            num nSigValue = 1
        pointRx pPointRx[2] = {x=490.110293, y=-600.305611, z=568.056156, rx=-6.599443, ry=-2.68541, rz=28.351195, shoulder=lefty, elbow=enegative, wrist=wpositive}
        string sID
      [48]
        bool bMarked
        jointRx jJointRx = {j1=-87.551314, j2=145.129335, j3=-83.085728, j4=182.11845, j5=63.691243, j6=-64.966658}
        pointRx pInter
        paraItem pParaItem
          [0]
            bool bSafePoint
            ifItem iIfItem
              [0]
                bool bANDOR[2]
                num nSigIndex[3]
                num nSigType[3]
                num nValue[3]
            mdesc mMdesc
            num nActionIndex = 42
            num nDelay
            num nMoveType = 1
            num nPercentage
            num nSigValue = 1
        pointRx pPointRx[2] = {x=61.349727, y=-652.129552, z=350.0734551, rx=-1.549449, ry=-1.96692, rz=28.421736, shoulder=lefty, elbow=enegative, wrist=wpositive}
        string sID
    string sID
  [Position6_point_blow]
    num nFrameIndex
    num nMoveID
    num nToolIndex
    pointItem pPointItem[64]
      [0]
        bool bMarked
        jointRx jJointRx
        pointRx pInter
        paraItem pParaItem
          [0]
            bool bSafePoint
            ifItem iIfItem
              [0]
                bool bANDOR[2]
                num nSigIndex[3]
                num nSigType[3]
                num nValue[3]
            mdesc mMdesc
            num nActionIndex = 43
            num nDelay
            num nMoveType = 4
            num nPercentage
            num nSigValue = 1
        pointRx pPointRx[2]
        string sID
      [1]
        bool bMarked
        jointRx jJointRx = {j1=-87.550712, j2=145.128314, j3=-83.0892365, j4=182.11811, j5=63.690987, j6=-64.966608}
        pointRx pInter
        paraItem pParaItem
          [0]
            bool bSafePoint
            ifItem iIfItem
              [0]
                bool bANDOR[2]
                num nSigIndex[3]
                num nSigType[3]
                num nValue[3]
            mdesc mMdesc
            num nActionIndex = 42
            num nDelay
            num nMoveType = 1
            num nPercentage
            num nSigValue = 1
        pointRx pPointRx[2] = {x=61.357264, y=-652.082, z=350.106484, rx=-1.553715, ry=-1.966811, rz=28.422241, shoulder=lefty, elbow=enegative, wrist=wpositive}
        string sID
      [2]
        bool bMarked
        jointRx jJointRx = {j1=-58.982134, j2=104.832128, j3=-61.565333, j4=183.343645, j5=42.668286, j6=-33.606181}
        pointRx pInter
        paraItem pParaItem
          [0]
            bool bSafePoint
            ifItem iIfItem
              [0]
                bool bANDOR[2]
                num nSigIndex[3]
                num nSigType[3]
                num nValue[3]
            mdesc mMdesc
            num nActionIndex = 42
            num nDelay
            num nMoveType = 1
            num nPercentage
            num nSigValue = 1
        pointRx pPointRx[2] = {x=416.397495, y=-633.838238, z=700.254781, rx=1.722211, ry=-1.608013, rz=89.88289, shoulder=lefty, elbow=enegative, wrist=wpositive}
        string sID
      [3]
        bool bMarked
        jointRx jJointRx = {j1=-62.332645, j2=107.50753, j3=-68.132801, j4=183.562396, j5=38.651057, j6=-30.577163}
        pointRx pInter
        paraItem pParaItem
          [0]
            bool bSafePoint
            ifItem iIfItem
              [0]
                bool bANDOR[2]
                num nSigIndex[3]
                num nSigType[3]
                num nValue[3]
            mdesc mMdesc
            num nActionIndex = 42
            num nDelay
            num nMoveType = 1
            num nPercentage
            num nSigValue = 1
        pointRx pPointRx[2] = {x=366.85786, y=-633.838275, z=700.254798, rx=1.721666, ry=-1.608681, rz=89.88277, shoulder=lefty, elbow=enegative, wrist=wpositive}
        string sID
      [4]
        bool bMarked
        jointRx jJointRx = {j1=-67.0327916, j2=110.2281, j3=-75.107293, j4=183.830258, j5=34.223084, j6=-26.259259}
        pointRx pInter
        paraItem pParaItem
          [0]
            bool bSafePoint
            ifItem iIfItem
              [0]
                bool bANDOR[2]
                num nSigIndex[3]
                num nSigType[3]
                num nValue[3]
            mdesc mMdesc
            num nActionIndex = 42
            num nDelay
            num nMoveType = 1
            num nPercentage
            num nSigValue = 1
        pointRx pPointRx[2] = {x=302.522929, y=-633.83826, z=700.254794, rx=1.721622, ry=-1.608914, rz=89.882692, shoulder=lefty, elbow=enegative, wrist=wpositive}
        string sID
      [5]
        bool bMarked
        jointRx jJointRx = {j1=-71.633736, j2=112.694899, j3=-81.788319, j4=184.160101, j5=29.845031, j6=-22.0972061}
        pointRx pInter
        paraItem pParaItem
          [0]
            bool bSafePoint
            ifItem iIfItem
              [0]
                bool bANDOR[2]
                num nSigIndex[3]
                num nSigType[3]
                num nValue[3]
            mdesc mMdesc
            num nActionIndex = 42
            num nDelay
            num nMoveType = 1
            num nPercentage
            num nSigValue = 1
        pointRx pPointRx[2] = {x=241.500206, y=-626.00943449, z=700.254792, rx=1.721289, ry=-1.608551, rz=89.882813, shoulder=lefty, elbow=enegative, wrist=wpositive}
        string sID
      [6]
        bool bMarked
        jointRx jJointRx = {j1=-65.27374, j2=114.413405, j3=-86.726434, j4=184.827216, j5=26.876761, j6=-29.158228}
        pointRx pInter
        paraItem pParaItem
          [0]
            bool bSafePoint
            ifItem iIfItem
              [0]
                bool bANDOR[2]
                num nSigIndex[3]
                num nSigType[3]
                num nValue[3]
            mdesc mMdesc
            num nActionIndex = 42
            num nDelay
            num nMoveType = 1
            num nPercentage
            num nSigValue = 1
        pointRx pPointRx[2] = {x=296.78184, y=-570.410131, z=700.254763, rx=1.722456, ry=-1.607129, rz=89.88308, shoulder=lefty, elbow=enegative, wrist=wpositive}
        string sID
      [7]
        bool bMarked
        jointRx jJointRx = {j1=-60.709616, j2=114.554511, j3=-87.145192, j4=184.986355, j5=26.782513, j6=-33.871303}
        pointRx pInter
        paraItem pParaItem
          [0]
            bool bSafePoint
            ifItem iIfItem
              [0]
                bool bANDOR[2]
                num nSigIndex[3]
                num nSigType[3]
                num nValue[3]
            mdesc mMdesc
            num nActionIndex = 42
            num nDelay
            num nMoveType = 1
            num nPercentage
            num nSigValue = 1
        pointRx pPointRx[2] = {x=338.875527, y=-541.934118, z=700.254791, rx=1.721113, ry=-1.608268, rz=89.882966, shoulder=lefty, elbow=enegative, wrist=wpositive}
        string sID
      [8]
        bool bMarked
        jointRx jJointRx = {j1=-66.643474, j2=118.657481, j3=-100.787497, j4=187.380827, j5=17.0599953, j6=-30.539636}
        pointRx pInter
        paraItem pParaItem
          [0]
            bool bSafePoint
            ifItem iIfItem
              [0]
                bool bANDOR[2]
                num nSigIndex[3]
                num nSigType[3]
                num nValue[3]
            mdesc mMdesc
            num nActionIndex = 42
            num nDelay
            num nMoveType = 1
            num nPercentage
            num nSigValue = 1
        pointRx pPointRx[2] = {x=251.241513, y=-503.208169, z=700.254788, rx=1.722301, ry=-1.608953, rz=89.882703, shoulder=lefty, elbow=enegative, wrist=wpositive}
        string sID
      [9]
        bool bMarked
        jointRx jJointRx = {j1=-65.0394334, j2=119.495527, j3=-104.191107, j4=188.704216, j5=14.582841, j6=-33.512784}
        pointRx pInter
        paraItem pParaItem
          [0]
            bool bSafePoint
            ifItem iIfItem
              [0]
                bool bANDOR[2]
                num nSigIndex[3]
                num nSigType[3]
                num nValue[3]
            mdesc mMdesc
            num nActionIndex = 42
            num nDelay
            num nMoveType = 1
            num nPercentage
            num nSigValue = 1
        pointRx pPointRx[2] = {x=255.846551, y=-476.313024, z=700.254767, rx=1.721654, ry=-1.607307, rz=89.883015, shoulder=lefty, elbow=enegative, wrist=wpositive}
        string sID
      [10]
        bool bMarked
        jointRx jJointRx = {j1=-71.0596735, j2=121.00750191, j3=-111.877772, j4=194.578806, j5=8.286602, j6=-33.494479}
        pointRx pInter
        paraItem pParaItem
          [0]
            bool bSafePoint
            ifItem iIfItem
              [0]
                bool bANDOR[2]
                num nSigIndex[3]
                num nSigType[3]
                num nValue[3]
            mdesc mMdesc
            num nActionIndex = 42
            num nDelay
            num nMoveType = 1
            num nPercentage
            num nSigValue = 1
        pointRx pPointRx[2] = {x=189.620191, y=-454.405925, z=700.254767, rx=1.721353, ry=-1.607377, rz=89.882905, shoulder=lefty, elbow=enegative, wrist=wpositive}
        string sID
      [11]
        bool bMarked
        jointRx jJointRx = {j1=-74.809464, j2=121.0382904, j3=-112.0769955, j4=194.59856, j5=7.974501, j6=-29.773551}
        pointRx pInter
        paraItem pParaItem
          [0]
            bool bSafePoint
            ifItem iIfItem
              [0]
                bool bANDOR[2]
                num nSigIndex[3]
                num nSigType[3]
                num nValue[3]
            mdesc mMdesc
            num nActionIndex = 42
            num nDelay
            num nMoveType = 1
            num nPercentage
            num nSigValue = 1
        pointRx pPointRx[2] = {x=160.082647, y=-465.491863, z=700.254784, rx=1.722803, ry=-1.608682, rz=89.882806, shoulder=lefty, elbow=enegative, wrist=wpositive}
        string sID
      [12]
        bool bMarked
        jointRx jJointRx = {j1=-76.815291, j2=120.680634, j3=-109.926019, j4=191.777648, j5=9.643692, j6=-24.919524}
        pointRx pInter
        paraItem pParaItem
          [0]
            bool bSafePoint
            ifItem iIfItem
              [0]
                bool bANDOR[2]
                num nSigIndex[3]
                num nSigType[3]
                num nValue[3]
            mdesc mMdesc
            num nActionIndex = 42
            num nDelay
            num nMoveType = 1
            num nPercentage
            num nSigValue = 1
        pointRx pPointRx[2] = {x=147.50556, y=-485.393693, z=700.254789, rx=1.722658, ry=-1.609045, rz=89.882735, shoulder=lefty, elbow=enegative, wrist=wpositive}
        string sID
      [13]
        bool bMarked
        jointRx jJointRx = {j1=-80.979539, j2=121.627826, j3=-116.887787, j4=209.4559, j5=3.779386, j6=-38.540773}
        pointRx pInter
        paraItem pParaItem
          [0]
            bool bSafePoint
            ifItem iIfItem
              [0]
                bool bANDOR[2]
                num nSigIndex[3]
                num nSigType[3]
                num nValue[3]
            mdesc mMdesc
            num nActionIndex = 42
            num nDelay
            num nMoveType = 1
            num nPercentage
            num nSigValue = 1
        pointRx pPointRx[2] = {x=105.438294, y=-448.641412, z=700.254346, rx=1.721348, ry=-1.60753, rz=89.882882, shoulder=lefty, elbow=enegative, wrist=wpositive}
        string sID
      [14]
        bool bMarked
        jointRx jJointRx = {j1=-97.0735787, j2=120.583034, j3=-109.386983, j4=169.0121648, j5=9.967554, j6=107.0502076}
        pointRx pInter
        paraItem pParaItem
          [0]
            bool bSafePoint
            ifItem iIfItem
              [0]
                bool bANDOR[2]
                num nSigIndex[3]
                num nSigType[3]
                num nValue[3]
            mdesc mMdesc
            num nActionIndex = 42
            num nDelay
            num nMoveType = 1
            num nPercentage
            num nSigValue = 1
        pointRx pPointRx[2] = {x=3.102788, y=-514.97816, z=700.254373, rx=1.629756, ry=1.702884, rz=179.149702, shoulder=lefty, elbow=enegative, wrist=wpositive}
        string sID
      [15]
        bool bMarked
        jointRx jJointRx = {j1=-98.785966, j2=121.589944, j3=-116.474742, j4=152.822693, j5=4.230949, j6=125.0509123}
        pointRx pInter
        paraItem pParaItem
          [0]
            bool bSafePoint
            ifItem iIfItem
              [0]
                bool bANDOR[2]
                num nSigIndex[3]
                num nSigType[3]
                num nValue[3]
            mdesc mMdesc
            num nActionIndex = 42
            num nDelay
            num nMoveType = 1
            num nPercentage
            num nSigValue = 1
        pointRx pPointRx[2] = {x=-4.455751, y=-466.481228, z=700.254288, rx=1.629056, ry=1.702249, rz=179.149669, shoulder=lefty, elbow=enegative, wrist=wpositive}
        string sID
      [16]
        bool bMarked
        jointRx jJointRx = {j1=-102.289362, j2=121.662055, j3=-117.287244, j4=147.396601, j5=3.732456, j6=133.989908}
        pointRx pInter
        paraItem pParaItem
          [0]
            bool bSafePoint
            ifItem iIfItem
              [0]
                bool bANDOR[2]
                num nSigIndex[3]
                num nSigType[3]
                num nValue[3]
            mdesc mMdesc
            num nActionIndex = 42
            num nDelay
            num nMoveType = 1
            num nPercentage
            num nSigValue = 1
        pointRx pPointRx[2] = {x=-30.830703, y=-458.833227, z=700.253116, rx=1.628925, ry=1.702444, rz=179.149706, shoulder=lefty, elbow=enegative, wrist=wpositive}
        string sID
      [17]
        bool bMarked
        jointRx jJointRx = {j1=-97.596795, j2=121.636094, j3=-116.996972, j4=154.0724475, j5=5.372504, j6=163.484863}
        pointRx pInter
        paraItem pParaItem
          [0]
            bool bSafePoint
            ifItem iIfItem
              [0]
                bool bANDOR[2]
                num nSigIndex[3]
                num nSigType[3]
                num nValue[3]
            mdesc mMdesc
            num nActionIndex = 42
            num nDelay
            num nMoveType = 1
            num nPercentage
            num nSigValue = 1
        pointRx pPointRx[2] = {x=11.0855283, y=-449.928798, z=700.263578, rx=0.116735, ry=2.351476, rz=-139.946822, shoulder=lefty, elbow=enegative, wrist=wpositive}
        string sID
      [18]
        bool bMarked
        jointRx jJointRx = {j1=-93.435678, j2=120.973902, j3=-111.67187, j4=165.758899, j5=9.616057, j6=147.540776}
        pointRx pInter
        paraItem pParaItem
          [0]
            bool bSafePoint
            ifItem iIfItem
              [0]
                bool bANDOR[2]
                num nSigIndex[3]
                num nSigType[3]
                num nValue[3]
            mdesc mMdesc
            num nActionIndex = 42
            num nDelay
            num nMoveType = 1
            num nPercentage
            num nSigValue = 1
        pointRx pPointRx[2] = {x=41.481677, y=-486.244692, z=700.26363, rx=0.117474, ry=2.35234, rz=-139.946783, shoulder=lefty, elbow=enegative, wrist=wpositive}
        string sID
      [19]
        bool bMarked
        jointRx jJointRx = {j1=-87.514361, j2=121.638618, j3=-117.0243701, j4=151.901605, j5=4.980778, j6=155.573887}
        pointRx pInter
        paraItem pParaItem
          [0]
            bool bSafePoint
            ifItem iIfItem
              [0]
                bool bANDOR[2]
                num nSigIndex[3]
                num nSigType[3]
                num nValue[3]
            mdesc mMdesc
            num nActionIndex = 42
            num nDelay
            num nMoveType = 1
            num nPercentage
            num nSigValue = 1
        pointRx pPointRx[2] = {x=89.805675, y=-444.448305, z=700.262762, rx=0.116151, ry=2.350833, rz=-139.946826, shoulder=lefty, elbow=enegative, wrist=wpositive}
        string sID
      [20]
        bool bMarked
        jointRx jJointRx = {j1=-85.538373, j2=121.159338, j3=-112.89672, j4=163.596021, j5=8.296682, j6=141.829296}
        pointRx pInter
        paraItem pParaItem
          [0]
            bool bSafePoint
            ifItem iIfItem
              [0]
                bool bANDOR[2]
                num nSigIndex[3]
                num nSigType[3]
                num nValue[3]
            mdesc mMdesc
            num nActionIndex = 42
            num nDelay
            num nMoveType = 1
            num nPercentage
            num nSigValue = 1
        pointRx pPointRx[2] = {x=107.297774, y=-470.450865, z=700.262819, rx=0.116544, ry=2.351714, rz=-139.94676, shoulder=lefty, elbow=enegative, wrist=wpositive}
        string sID
      [21]
        bool bMarked
        jointRx jJointRx = {j1=-80.389938, j2=121.305327, j3=-113.961147, j4=161.375696, j5=7.211507, j6=138.92232}
        pointRx pInter
        paraItem pParaItem
          [0]
            bool bSafePoint
            ifItem iIfItem
              [0]
                bool bANDOR[2]
                num nSigIndex[3]
                num nSigType[3]
                num nValue[3]
            mdesc mMdesc
            num nActionIndex = 42
            num nDelay
            num nMoveType = 1
            num nPercentage
            num nSigValue = 1
        pointRx pPointRx[2] = {x=147.836969, y=-453.554332, z=700.262491, rx=0.115759, ry=2.349936, rz=-139.946858, shoulder=lefty, elbow=enegative, wrist=wpositive}
        string sID
      [22]
        bool bMarked
        jointRx jJointRx = {j1=-74.160542, j2=121.48868, j3=-115.480429, j4=163.296331, j5=4.15176, j6=89.975533}
        pointRx pInter
        paraItem pParaItem
          [0]
            bool bSafePoint
            ifItem iIfItem
              [0]
                bool bANDOR[2]
                num nSigIndex[3]
                num nSigType[3]
                num nValue[3]
            mdesc mMdesc
            num nActionIndex = 42
            num nDelay
            num nMoveType = 1
            num nPercentage
            num nSigValue = 1
        pointRx pPointRx[2] = {x=187.654652, y=-440.110471, z=700.252779, rx=1.628669, ry=1.701382, rz=179.149675, shoulder=lefty, elbow=enegative, wrist=wpositive}
        string sID
      [23]
        bool bMarked
        jointRx jJointRx = {j1=-69.509661, j2=119.265921, j3=-103.220112, j4=175.749132, j5=13.961301, j6=72.790426}
        pointRx pInter
        paraItem pParaItem
          [0]
            bool bSafePoint
            ifItem iIfItem
              [0]
                bool bANDOR[2]
                num nSigIndex[3]
                num nSigType[3]
                num nValue[3]
            mdesc mMdesc
            num nActionIndex = 42
            num nDelay
            num nMoveType = 1
            num nPercentage
            num nSigValue = 1
        pointRx pPointRx[2] = {x=250.0960558, y=-500.875002, z=700.252775, rx=1.628687, ry=1.702386, rz=179.149806, shoulder=lefty, elbow=enegative, wrist=wpositive}
        string sID
      [24]
        bool bMarked
        jointRx jJointRx = {j1=-65.451313, j2=120.0346612, j3=-106.615882, j4=175.540521, j5=11.264344, j6=68.982362}
        pointRx pInter
        paraItem pParaItem
          [0]
            bool bSafePoint
            ifItem iIfItem
              [0]
                bool bANDOR[2]
                num nSigIndex[3]
                num nSigType[3]
                num nValue[3]
            mdesc mMdesc
            num nActionIndex = 42
            num nDelay
            num nMoveType = 1
            num nPercentage
            num nSigValue = 1
        pointRx pPointRx[2] = {x=274.930404, y=-463.298611, z=700.25277, rx=1.6286, ry=1.700384, rz=179.149585, shoulder=lefty, elbow=enegative, wrist=wpositive}
        string sID
      [25]
        bool bMarked
        jointRx jJointRx = {j1=-63.0913911, j2=120.463088, j3=-108.745441, j4=175.274971, j5=9.527094, j6=66.910352}
        pointRx pInter
        paraItem pParaItem
          [0]
            bool bSafePoint
            ifItem iIfItem
              [0]
                bool bANDOR[2]
                num nSigIndex[3]
                num nSigType[3]
                num nValue[3]
            mdesc mMdesc
            num nActionIndex = 42
            num nDelay
            num nMoveType = 1
            num nPercentage
            num nSigValue = 1
        pointRx pPointRx[2] = {x=286.920288, y=-439.796835, z=700.252783, rx=1.628449, ry=1.702261, rz=179.149771, shoulder=lefty, elbow=enegative, wrist=wpositive}
        string sID
      [26]
        bool bMarked
        jointRx jJointRx = {j1=-60.107122, j2=120.743514, j3=-110.280684, j4=175.353325, j5=8.229554, j6=63.86699}
        pointRx pInter
        paraItem pParaItem
          [0]
            bool bSafePoint
            ifItem iIfItem
              [0]
                bool bANDOR[2]
                num nSigIndex[3]
                num nSigType[3]
                num nValue[3]
            mdesc mMdesc
            num nActionIndex = 42
            num nDelay
            num nMoveType = 1
            num nPercentage
            num nSigValue = 1
        pointRx pPointRx[2] = {x=303.628134, y=-416.218815, z=700.252788, rx=1.628466, ry=1.702202, rz=179.149747, shoulder=lefty, elbow=enegative, wrist=wpositive}
        string sID
      [27]
        bool bMarked
        jointRx jJointRx = {j1=-63.992151, j2=118.544695, j3=-100.353777, j4=177.0428516, j5=16.00047448, j6=65.992969}
        pointRx pInter
        paraItem pParaItem
          [0]
            bool bSafePoint
            ifItem iIfItem
              [0]
                bool bANDOR[2]
                num nSigIndex[3]
                num nSigType[3]
                num nValue[3]
            mdesc mMdesc
            num nActionIndex = 42
            num nDelay
            num nMoveType = 1
            num nPercentage
            num nSigValue = 1
        pointRx pPointRx[2] = {x=303.593559, y=-492.00120121, z=700.25275, rx=1.629773, ry=1.701529, rz=179.149557, shoulder=lefty, elbow=enegative, wrist=wpositive}
        string sID
      [28]
        bool bMarked
        jointRx jJointRx = {j1=-65.604658, j2=115.34522, j3=-89.535997, j4=177.811149, j5=23.638027, j6=66.767236}
        pointRx pInter
        paraItem pParaItem
          [0]
            bool bSafePoint
            ifItem iIfItem
              [0]
                bool bANDOR[2]
                num nSigIndex[3]
                num nSigType[3]
                num nValue[3]
            mdesc mMdesc
            num nActionIndex = 42
            num nDelay
            num nMoveType = 1
            num nPercentage
            num nSigValue = 1
        pointRx pPointRx[2] = {x=316.105522, y=-557.406438, z=700.252765, rx=1.629152, ry=1.702122, rz=179.149764, shoulder=lefty, elbow=enegative, wrist=wpositive}
        string sID
      [29]
        bool bMarked
        jointRx jJointRx = {j1=-68.955824, j2=108.932967, j3=-71.74331, j4=178.253914, j5=35.0703752, j6=69.540198}
        pointRx pInter
        paraItem pParaItem
          [0]
            bool bSafePoint
            ifItem iIfItem
              [0]
                bool bANDOR[2]
                num nSigIndex[3]
                num nSigType[3]
                num nValue[3]
            mdesc mMdesc
            num nActionIndex = 42
            num nDelay
            num nMoveType = 1
            num nPercentage
            num nSigValue = 1
        pointRx pPointRx[2] = {x=316.0702808, y=-657.877777, z=700.252731, rx=1.629581, ry=1.701668, rz=179.149612, shoulder=lefty, elbow=enegative, wrist=wpositive}
        string sID
      [30]
        bool bMarked
        jointRx jJointRx = {j1=-63.428303, j2=105.599126, j3=-63.42748, j4=178.764025, j5=39.960548, j6=63.523315}
        pointRx pInter
        paraItem pParaItem
          [0]
            bool bSafePoint
            ifItem iIfItem
              [0]
                bool bANDOR[2]
                num nSigIndex[3]
                num nSigType[3]
                num nValue[3]
            mdesc mMdesc
            num nActionIndex = 42
            num nDelay
            num nMoveType = 1
            num nPercentage
            num nSigValue = 1
        pointRx pPointRx[2] = {x=392.672125, y=-657.853849, z=700.276087, rx=1.628612, ry=1.701821, rz=179.138765, shoulder=lefty, elbow=enegative, wrist=wpositive}
        string sID
      [31]
        bool bMarked
        jointRx jJointRx = {j1=-64.321332, j2=88.690196, j3=-45.113442, j4=178.747654, j5=41.378269, j6=64.407958}
        pointRx pInter
        paraItem pParaItem
          [0]
            bool bSafePoint
            ifItem iIfItem
              [0]
                bool bANDOR[2]
                num nSigIndex[3]
                num nSigType[3]
                num nValue[3]
            mdesc mMdesc
            num nActionIndex = 42
            num nDelay
            num nMoveType = 1
            num nPercentage
            num nSigValue = 1
        pointRx pPointRx[2] = {x=392.636913, y=-684.559631, z=817.184286, rx=1.629027, ry=1.701529, rz=179.138589, shoulder=lefty, elbow=enegative, wrist=wpositive}
        string sID
      [32]
        bool bMarked
        jointRx jJointRx = {j1=-64.968443, j2=76.908071, j3=-27.68217, j4=178.834761, j5=47.0360379, j6=64.909112}
        pointRx pInter
        paraItem pParaItem
          [0]
            bool bSafePoint
            ifItem iIfItem
              [0]
                bool bANDOR[2]
                num nSigIndex[3]
                num nSigType[3]
                num nValue[3]
            mdesc mMdesc
            num nActionIndex = 42
            num nDelay
            num nMoveType = 1
            num nPercentage
            num nSigValue = 1
        pointRx pPointRx[2] = {x=392.63674, y=-705.0468714, z=873.404329, rx=1.628998, ry=1.701548, rz=179.138605, shoulder=lefty, elbow=enegative, wrist=wpositive}
        string sID
      [33]
        bool bMarked
        jointRx jJointRx = {j1=-62.336449, j2=89.481455, j3=-54.547425, j4=178.610325, j5=32.711346, j6=62.654003}
        pointRx pInter
        paraItem pParaItem
          [0]
            bool bSafePoint
            ifItem iIfItem
              [0]
                bool bANDOR[2]
                num nSigIndex[3]
                num nSigType[3]
                num nValue[3]
            mdesc mMdesc
            num nActionIndex = 42
            num nDelay
            num nMoveType = 1
            num nPercentage
            num nSigValue = 1
        pointRx pPointRx[2] = {x=392.637106, y=-627.212597, z=851.844705, rx=1.627027, ry=1.700481, rz=179.138679, shoulder=lefty, elbow=enegative, wrist=wpositive}
        string sID
      [34]
        bool bMarked
        jointRx jJointRx = {j1=-60.214263, j2=94.794241, j3=-66.773415, j4=178.463697, j5=25.772301, j6=60.747514}
        pointRx pInter
        paraItem pParaItem
          [0]
            bool bSafePoint
            ifItem iIfItem
              [0]
                bool bANDOR[2]
                num nSigIndex[3]
                num nSigType[3]
                num nValue[3]
            mdesc mMdesc
            num nActionIndex = 42
            num nDelay
            num nMoveType = 1
            num nPercentage
            num nSigValue = 1
        pointRx pPointRx[2] = {x=392.637091, y=-573.593172, z=839.237969, rx=1.626982, ry=1.700524, rz=179.13871, shoulder=lefty, elbow=enegative, wrist=wpositive}
        string sID
      [35]
        bool bMarked
        jointRx jJointRx = {j1=-55.995459, j2=94.871223, j3=-77.350718, j4=178.0932115, j5=15.228667, j6=56.988296}
        pointRx pInter
        paraItem pParaItem
          [0]
            bool bSafePoint
            ifItem iIfItem
              [0]
                bool bANDOR[2]
                num nSigIndex[3]
                num nSigType[3]
                num nValue[3]
            mdesc mMdesc
            num nActionIndex = 42
            num nDelay
            num nMoveType = 1
            num nPercentage
            num nSigValue = 1
        pointRx pPointRx[2] = {x=392.637078, y=-484.790879, z=868.772586, rx=1.626877, ry=1.701216, rz=179.138854, shoulder=lefty, elbow=enegative, wrist=wpositive}
        string sID
      [36]
        bool bMarked
        jointRx jJointRx = {j1=-58.229299, j2=114.285829, j3=-86.304494, j4=178.642261, j5=25.707127, j6=58.603666}
        pointRx pInter
        paraItem pParaItem
          [0]
            bool bSafePoint
            ifItem iIfItem
              [0]
                bool bANDOR[2]
                num nSigIndex[3]
                num nSigType[3]
                num nValue[3]
            mdesc mMdesc
            num nActionIndex = 42
            num nDelay
            num nMoveType = 1
            num nPercentage
            num nSigValue = 1
        pointRx pPointRx[2] = {x=392.637007, y=-529.258957, z=700.0975269, rx=1.629049, ry=1.701252, rz=179.138503, shoulder=lefty, elbow=enegative, wrist=wpositive}
        string sID
      [37]
        bool bMarked
        jointRx jJointRx = {j1=-82.703196, j2=116.122044, j3=-91.853722, j4=179.533458, j5=22.561363, j6=-8.781235}
        pointRx pInter
        paraItem pParaItem
          [0]
            bool bSafePoint
            ifItem iIfItem
              [0]
                bool bANDOR[2]
                num nSigIndex[3]
                num nSigType[3]
                num nValue[3]
            mdesc mMdesc
            num nActionIndex = 42
            num nDelay
            num nMoveType = 1
            num nPercentage
            num nSigValue = 1
        pointRx pPointRx[2] = {x=130.0386713, y=-609.589422, z=700.0975633, rx=1.671086, ry=0.394403, rz=88.0816451, shoulder=lefty, elbow=enegative, wrist=wpositive}
        string sID
      [38]
        bool bMarked
        jointRx jJointRx = {j1=-82.0614145, j2=118.602251, j3=-100.420616, j4=179.303357, j5=16.477589, j6=-7.920976}
        pointRx pInter
        paraItem pParaItem
          [0]
            bool bSafePoint
            ifItem iIfItem
              [0]
                bool bANDOR[2]
                num nSigIndex[3]
                num nSigType[3]
                num nValue[3]
            mdesc mMdesc
            num nActionIndex = 42
            num nDelay
            num nMoveType = 1
            num nPercentage
            num nSigValue = 1
        pointRx pPointRx[2] = {x=130.0386769, y=-558.013851, z=700.0975609, rx=1.661587, ry=0.431173, rz=89.346263, shoulder=lefty, elbow=enegative, wrist=wpositive}
        string sID
      [39]
        bool bMarked
        jointRx jJointRx = {j1=-90.0104561, j2=120.70672, j3=-109.816065, j4=177.317534, j5=9.238811, j6=2.005015}
        pointRx pInter
        paraItem pParaItem
          [0]
            bool bSafePoint
            ifItem iIfItem
              [0]
                bool bANDOR[2]
                num nSigIndex[3]
                num nSigType[3]
                num nValue[3]
            mdesc mMdesc
            num nActionIndex = 42
            num nDelay
            num nMoveType = 1
            num nPercentage
            num nSigValue = 1
        pointRx pPointRx[2] = {x=53.663817, y=-510.218495, z=700.0975573, rx=1.661871, ry=0.430213, rz=89.346845, shoulder=lefty, elbow=enegative, wrist=wpositive}
        string sID
      [40]
        bool bMarked
        jointRx jJointRx = {j1=-98.300868, j2=121.852736, j3=-119.389976, j4=142.928524, j5=1.104688, j6=44.711227}
        pointRx pInter
        paraItem pParaItem
          [0]
            bool bSafePoint
            ifItem iIfItem
              [0]
                bool bANDOR[2]
                num nSigIndex[3]
                num nSigType[3]
                num nValue[3]
            mdesc mMdesc
            num nActionIndex = 42
            num nDelay
            num nMoveType = 1
            num nPercentage
            num nSigValue = 1
        pointRx pPointRx[2] = {x=-8.738518, y=-446.473036, z=700.0947095, rx=1.660849, ry=0.430654, rz=89.346953, shoulder=lefty, elbow=enegative, wrist=wpositive}
        string sID
      [41]
        bool bMarked
        jointRx jJointRx = {j1=-101.944431, j2=121.840245, j3=-119.156799, j4=146.219817, j5=1.37852, j6=45.0598803}
        pointRx pInter
        paraItem pParaItem
          [0]
            bool bSafePoint
            ifItem iIfItem
              [0]
                bool bANDOR[2]
                num nSigIndex[3]
                num nSigType[3]
                num nValue[3]
            mdesc mMdesc
            num nActionIndex = 42
            num nDelay
            num nMoveType = 1
            num nPercentage
            num nSigValue = 1
        pointRx pPointRx[2] = {x=-36.505296, y=-446.471107, z=700.0993486, rx=1.662873, ry=0.431649, rz=89.346951, shoulder=lefty, elbow=enegative, wrist=wpositive}
        string sID
      [42]
        bool bMarked
        jointRx jJointRx = {j1=-83.477862, j2=120.163104, j3=-107.0210872, j4=187.573096, j5=13.00753743, j6=-104.399477}
        pointRx pInter
        paraItem pParaItem
          [0]
            bool bSafePoint
            ifItem iIfItem
              [0]
                bool bANDOR[2]
                num nSigIndex[3]
                num nSigType[3]
                num nValue[3]
            mdesc mMdesc
            num nActionIndex = 42
            num nDelay
            num nMoveType = 1
            num nPercentage
            num nSigValue = 1
        pointRx pPointRx[2] = {x=93.575962, y=-508.878606, z=700.0975715, rx=0.435679, ry=-1.661103, rz=-0.4937, shoulder=lefty, elbow=enegative, wrist=wpositive}
        string sID
      [43]
        bool bMarked
        jointRx jJointRx = {j1=-82.561979, j2=121.615974, j3=-116.238306, j4=198.28183, j5=5.43426, j6=-116.137422}
        pointRx pInter
        paraItem pParaItem
          [0]
            bool bSafePoint
            ifItem iIfItem
              [0]
                bool bANDOR[2]
                num nSigIndex[3]
                num nSigType[3]
                num nValue[3]
            mdesc mMdesc
            num nActionIndex = 42
            num nDelay
            num nMoveType = 1
            num nPercentage
            num nSigValue = 1
        pointRx pPointRx[2] = {x=93.575581, y=-445.271705, z=700.110228, rx=0.4348, ry=-1.660062, rz=-0.491221, shoulder=lefty, elbow=enegative, wrist=wpositive}
        string sID
      [44]
        bool bMarked
        jointRx jJointRx = {j1=-81.917883, j2=121.906713, j3=-121.128234, j4=251.166903, j5=1.801978, j6=-169.734998}
        pointRx pInter
        paraItem pParaItem
          [0]
            bool bSafePoint
            ifItem iIfItem
              [0]
                bool bANDOR[2]
                num nSigIndex[3]
                num nSigType[3]
                num nValue[3]
            mdesc mMdesc
